(*
	Posts each accepted batch as one OTLP/HTTP ProtoJSON TracesData request to an OTLP
	collector, for example 'http://192.168.1.10:4318/v1/traces'. Call the instance, or tick,
	every scan: the exporter is busy from export until currentState reaches done or error.
	The batch is released at either end, and an error is reported by tick until the next
	batch is accepted. A response outside 2xx is an error; nothing is retried.
*)
FUNCTION_BLOCK FB_SpanExporter_HTTP EXTENDS FB_SpanExporter_Base
VAR_OUTPUT
	currentState: E_HttpExporterState;
	statusCode: UINT;  // the HTTP status code received for the last completed request
END_VAR

VAR
	_execute: BOOL;
	_urlParsed: BOOL;
	_endpoint: ST_HttpEndpoint;
	_len: UDINT;
	_execRTrig: R_TRIG;
	_pString: POINTER TO STRING;
	_jsonVal: SJsonValue;
	_computedState: E_HttpExporterState;
	_failureReason: E_SpanExporterFailureReason;
	_serializationFailureReason: E_ProtoJsonSerializerFailureReason;
	_serializer: FB_SpanProtoJsonSerializer;
	_client: FB_IotHttpClient;
	_request: FB_IotHttpRequest;
	_header: FB_IotHttpHeaderFieldMap;
END_VAR

THIS^.tick(failureReason=>THIS^._callFailureReason);

METHOD export: BOOL
VAR_IN_OUT
	spans: FB_SpanQueue;
END_VAR
VAR_INPUT
	count: UDINT;
END_VAR
VAR_OUTPUT
	failureReason: E_SpanExporterFailureReason;
END_VAR
// a finished exporter accepts the next batch at once
IF THIS^.currentState = E_HttpExporterState.done OR THIS^.currentState = E_HttpExporterState.error THEN
	THIS^.currentState := E_HttpExporterState.idle;
	THIS^._computedState := E_HttpExporterState.idle;
END_IF
export := SUPER^.export(
	spans:=spans,
	count:=count,
	failureReason=>failureReason
);
IF export THEN
	THIS^._failureReason := E_SpanExporterFailureReason.NA;
	THIS^._serializationFailureReason := E_ProtoJsonSerializerFailureReason.NA;
END_IF
END_METHOD

(*
	Releases a payload buffer that is still in flight. The FB_IotHttpRequest reading it is
	destroyed with this instance, so nothing uses the buffer afterwards. TwinCAT then
	runs FB_SpanExporter_Base.FB_Exit, which releases the accepted spans.
*)
METHOD FB_Exit : BOOL
VAR_INPUT
	bInCopyCode: BOOL;  // TRUE: the instance is being copied during an online change
END_VAR
// during an online change the copy keeps the buffer, so it must not be released here
IF NOT bInCopyCode AND _pString <> 0 THEN
	__DELETE(_pString);
	_pString := 0;
END_IF
END_METHOD

METHOD FB_Init: BOOL
VAR_INPUT
	bInitRetains: BOOL; // TRUE: the retain variables are initialized (reset warm / reset cold)
	bInCopyCode: BOOL;  // TRUE: the instance will be copied to the copy code afterward (online change)
	url: T_MaxString;  // full endpoint URL, e.g. 'http://192.168.1.10:4318/v1/traces'
	bNoServerCertCheck: BOOL := FALSE;  // allow HTTPS connections to servers with self-signed certificates
END_VAR
THIS^.currentState := E_HttpExporterState.idle;
THIS^._computedState := E_HttpExporterState.idle;

THIS^._urlParsed := F_ParseHttpUrl(url:=url, endpoint=>THIS^._endpoint);

THIS^._client.sHostName := THIS^._endpoint.host;
THIS^._client.nHostPort := THIS^._endpoint.port;
THIS^._client.bKeepAlive := TRUE;
THIS^._client.tConnectionTimeout := T#10S;
IF THIS^._endpoint.useTls THEN
	THIS^._client.stTLS.bNoServerCertCheck := bNoServerCertCheck;
END_IF

THIS^._request.sContentType := 'application/json';
END_METHOD

METHOD isBusy : BOOL
isBusy := THIS^._exportActive;
END_METHOD

METHOD tick : BOOL
VAR_OUTPUT
	failureReason: E_SpanExporterFailureReason;
END_VAR
tick := TRUE;
failureReason := E_SpanExporterFailureReason.NA;

_execute := THIS^._exportActive;
_execRTrig(CLK := _execute AND_THEN THIS^._spans.count > 0);

CASE currentState OF
	E_HttpExporterState.idle:
		IF _execRTrig.Q THEN
			_failureReason := E_SpanExporterFailureReason.NA;
			_serializationFailureReason := E_ProtoJsonSerializerFailureReason.NA;
			IF NOT THIS^._urlParsed THEN
				_failureReason := E_SpanExporterFailureReason.HTTP_URL_PARSE_FAILURE;
				_computedState := E_HttpExporterState.error;
			ELSE
				_computedState := E_HttpExporterState.serializing;
			END_IF
		END_IF

	E_HttpExporterState.serializing:
		// the serializer drains the batch; buffer the TracesData document as the payload
		IF NOT _serializer.serializeTracesData(
			spans:=THIS^._spans,
			failureReason=>_serializationFailureReason
		) THEN
			_failureReason := E_SpanExporterFailureReason.SERIALIZATION_FAILURE;
			_computedState := E_HttpExporterState.error;
		ELSE
			_jsonVal := _serializer.jsonValue;
			IF _jsonVal = 0 OR_ELSE NOT _serializer.parser.IsObject(_jsonVal) THEN
				_failureReason := E_SpanExporterFailureReason.SERIALIZATION_FAILURE;
				_computedState := E_HttpExporterState.error;
			ELSE
				_len := _serializer.parser.GetJsonLength(_jsonVal);  // includes the null terminating character
				IF _len = 0 THEN
					_failureReason := E_SpanExporterFailureReason.SERIALIZATION_FAILURE;
					_computedState := E_HttpExporterState.error;
				ELSE
					_pString := __NEW(BYTE, _len);
					IF _pString = 0 THEN
						_failureReason := E_SpanExporterFailureReason.BUFFER_ALLOCATION_FAILURE;
						_computedState := E_HttpExporterState.error;
					ELSE
						_serializer.parser.CopyJson(_jsonVal, _pString^, _len);
						_computedState := E_HttpExporterState.sending;
					END_IF
				END_IF
			END_IF
		END_IF

	E_HttpExporterState.sending:
		IF NOT _request.bBusy THEN
			IF _request.SendRequest(
				sUri := THIS^._endpoint.path,
				fbClient := THIS^._client,
				eRequestType := ETcIotHttpRequestType.HTTP_POST,
				pContent := _pString,
				nContentSize := _len - 1,
				fbHeader := THIS^._header
			) THEN
				_computedState := E_HttpExporterState.waiting;
			ELSE
				IF _pString <> 0 THEN __DELETE(_pString); _pString := 0; END_IF
				_failureReason := E_SpanExporterFailureReason.HTTP_REQUEST_FAILURE;
				_computedState := E_HttpExporterState.error;
			END_IF
		END_IF

	E_HttpExporterState.waiting:
		IF NOT _request.bBusy THEN
			_computedState := E_HttpExporterState.processing;
		END_IF

	E_HttpExporterState.processing:
		IF _request.bError THEN
			IF _pString <> 0 THEN __DELETE(_pString); _pString := 0; END_IF
			_failureReason := E_SpanExporterFailureReason.HTTP_REQUEST_FAILURE;
			_computedState := E_HttpExporterState.error;
		ELSE
			statusCode := _request.nStatusCode;
			IF statusCode < 200 OR_ELSE statusCode >= 300 THEN
				IF _pString <> 0 THEN __DELETE(_pString); _pString := 0; END_IF
				_failureReason := E_SpanExporterFailureReason.HTTP_STATUS_FAILURE;
				_computedState := E_HttpExporterState.error;
			ELSE
				IF _pString <> 0 THEN __DELETE(_pString); _pString := 0; END_IF
				_computedState := E_HttpExporterState.done;
			END_IF
		END_IF

	E_HttpExporterState.done:
		IF NOT _execute THEN
			_computedState := E_HttpExporterState.idle;
		END_IF

	E_HttpExporterState.error:
		// keep the failure until export accepts a new batch
END_CASE

currentState := _computedState;

IF currentState = E_HttpExporterState.done
	OR_ELSE currentState = E_HttpExporterState.error THEN
	THIS^.free();
END_IF

THIS^._client.Execute();

IF currentState = E_HttpExporterState.error THEN
	tick := FALSE;
	failureReason := _failureReason;
END_IF
END_METHOD

END_FUNCTION_BLOCK

(* stored: Version 1.1.0.1
   POU FB_SpanExporter_HTTP: Id {f345cdfb-17a2-41e9-81c9-d9480cfbb5ea}, SpecialFunc None
   Method export: Id {23053720-09e7-4425-9a75-b490ecc94e69}
   Method FB_Exit: Id {f72f4f48-02e2-4781-ac1d-f0952810c37e}
   Method FB_Init: Id {8924758c-3494-4d4e-ac99-0029f9c87ef7}
   Method isBusy: Id {3c56e687-e28a-4636-8917-4eb786e5a97e}
   Method tick: Id {6d675a02-42e2-454b-b95a-21e2bdb2a3a6} *)
